// TIA Portal V20 export
TYPE "WT2_Pf_Befehl_UDT"
   STRUCT
      iHandshake : Int;
      Datum : Array[0..9] of Char;
      Zeit : Array[0..7] of Char;
      byKonfigSetFix : Byte;
      bySammelquit : Byte;
      byKonfigSetZykl : Byte;
      by23_Reserve : Byte;
      byReserve : Array[0..39] of Byte;
   END_STRUCT;
END_TYPE
